Fanuc KAREL source: KA00221.KL

PROGRAM KA00221
%NOLOCKGROUP
VAR
  SRC: ARRAY[4] OF JOINTPOS
  DST: ARRAY[4] OF BYTE
BEGIN
  DST = SRC
END KA00221
